Fanuc KAREL source: KO00149.KL

PROGRAM KO00149
%NOLOCKGROUP
VAR
  R: REAL
  CFG: CONFIG
  OUT: XYZWPR
  N: INTEGER
BEGIN
  N = 1
  R = 2.0
  CFG.CFG_FLIP = TRUE
  OUT = POS(R, R, R, R, R, N, CFG)
END KO00149
